(* PLC project zarechnaya.project, CODESYS CODESYS V3.5 SP17 Patch 3 *)
(* stored: creationDateTime 2026-10-20T05:42:22.1846158, modificationDateTime 1601-01-01T03:00:00 *)

(* FB_Latch — фиксация команд пульта фильтра (ST, FUNCTION_BLOCK). Поведение (модель scenarios/reference/model_FB_Latch.py): - xSr — SR(SET1 := xSet, RESET := xReset): установка доминирует, при SET = RESET = 1 → TRUE; - xRs — RS(SET := xSet, RESET1 := xReset): сброс доминирует, при SET = RESET = 1 → FALSE (одноимённые блоки S7 — наоборот: C2S7-SEM-SRRS, CDS_SR/CDS_RS); - CTU(CU := xCu, RESET := xReset, PV := 3): wCu — счёт фронтов, xCuQ — wCu ≥ 3; RESET обнуляет; - CTD(CD := xCd, LOAD := xLoad, PV := 2): LOAD ставит 2, фронт CD уменьшает до 0 и не ниже, xCdQ — wCd = 0 (WORD без знака: стоит на нуле; проба M0); - xRise/xFall — R_TRIG/F_TRIG по xClk; F_TRIG на первом вызове с CLK = FALSE спада не даёт (M0). *)
FUNCTION_BLOCK FB_Latch
  VAR_INPUT
    xSet : BOOL;
    xReset : BOOL;
    xCu : BOOL;
    xCd : BOOL;
    xLoad : BOOL;
    xClk : BOOL;
  END_VAR
  VAR_OUTPUT
    xSr : BOOL;
    xRs : BOOL;
    xCuQ : BOOL;
    xCdQ : BOOL;
    wCu : WORD;
    wCd : WORD;
    xRise : BOOL;
    xFall : BOOL;
  END_VAR
  VAR
    fbSr : SR;
    fbRs : RS;
    fbCtu : CTU;
    fbCtd : CTD;
    fbRise : R_TRIG;
    fbFall : F_TRIG;
  END_VAR

            fbSr(SET1 := xSet, RESET := xReset, Q1 => xSr);
fbRs(SET := xSet, RESET1 := xReset, Q1 => xRs);
fbCtu(CU := xCu, RESET := xReset, PV := 3, Q => xCuQ, CV => wCu);
fbCtd(CD := xCd, LOAD := xLoad, PV := 2, Q => xCdQ, CV => wCd);
fbRise(CLK := xClk, Q => xRise);
fbFall(CLK := xClk, Q => xFall);

          
END_FUNCTION_BLOCK
